FUNCTION_BLOCK EjectorCtrl (* Basic Function Block Type *)
  (* Standard: 61499-2 *)
  (* Version 0.0, 7/2/2026, Template *)
  PACKAGE Main;
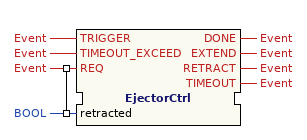
  EVENT_INPUT
    TRIGGER; (* Initialization Request *)
    TIMEOUT_EXCEED;
    REQ WITH retracted; (* Normal Execution Request *)
  END_EVENT
  EVENT_OUTPUT
    DONE; (* Initialization Confirm *)
    EXTEND; (* Execution Confirmation *)
    RETRACT;
    TIMEOUT;
  END_EVENT
  VAR_INPUT
    retracted : BOOL; (* Input event qualifier *)
  END_VAR
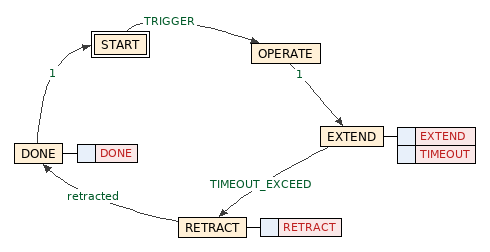
  EC_STATES
    START; (* Initial State *)
    OPERATE;
    EXTEND : -> EXTEND, -> TIMEOUT;
    RETRACT : -> RETRACT;
    DONE : -> DONE;
  END_STATES
  EC_TRANSITIONS
    START TO OPERATE := TRIGGER;
    OPERATE TO EXTEND := 1;
    EXTEND TO RETRACT := TIMEOUT_EXCEED;
    RETRACT TO DONE := retracted;
    DONE TO START := 1;
  END_TRANSITIONS
  ALGORITHM INIT IN ST: (* Initialization algorithm *)
;
  END_ALGORITHM
  ALGORITHM REQ IN ST: (* Normally executed algorithm *)
;
  END_ALGORITHM
END_FUNCTION_BLOCK
